// TIA Portal project "EXERCICE_IHM" (V16)

(* hardware
DEVICE "HMI_1"  KTP700 Basic PN
   slot 0: "HMI_1"  KTP700 Basic PN  6AV2 123-2GB03-0AX0  16.0.0.0
   slot 1: "HMI_RT_1"  KTP700 Basic PN  6AV2 123-2GB03-0AX0  16.0.0.0
   slot 5: "HMI_1.IE_CP_1"  PROFINET Interface  16.0.0.0
      slot 1: "Interface PROFINET_1"  PROFINET Interface
         slot 1: "Port_1"  Port
DEVICE "Station S7-1200_1"  S7-1200 Station
   slot 0: "Châssis_0"  S7-1200 Rack  Rack  V1.0
   slot 1: "PLC_1"  CPU 1214C AC/DC/Rly  6ES7 214-1BG40-0XB0  V4.4
*)

// ===== PLC "PLC_1"  CPU 1214C AC/DC/Rly =====

VAR_GLOBAL   // PLC tag table "Table de variables standard"
   "START" AT %I0.0 : Bool;
   "STOP" AT %I0.1 : Bool;
   "Moteur" AT %Q0.0 : Bool;
   "H1" AT %Q0.1 : Bool;
   "Clock_Byte" AT %MB0 : Byte;
   "Clock_10Hz" AT %M0.0 : Bool;
   "Clock_5Hz" AT %M0.1 : Bool;
   "Clock_2.5Hz" AT %M0.2 : Bool;
   "Clock_2Hz" AT %M0.3 : Bool;
   "Clock_1.25Hz" AT %M0.4 : Bool;
   "Clock_1Hz" AT %M0.5 : Bool;
   "Clock_0.625Hz" AT %M0.6 : Bool;
   "Clock_0.5Hz" AT %M0.7 : Bool;
   "HMI VENTILATEUR" AT %Q0.2 : Bool;
   "VENTILATEUR" AT %Q0.3 : Bool;
   "HMI MEMEUR" AT %Q0.4 : Bool;
END_VAR

ORGANIZATION_BLOCK "Main"   // OB1, LAD, ProgramCycle
TITLE = "Main Program Sweep (Cycle)"
{ S7_Optimized_Access := 'TRUE' }
VERSION : 0.1
   VAR_INPUT
      Initial_Call : Bool;   // Initial call of this OB
      Remanence : Bool;   // =True, if remanent data are available
   END_VAR
BEGIN

REGION Network 1
   // MOTEUR
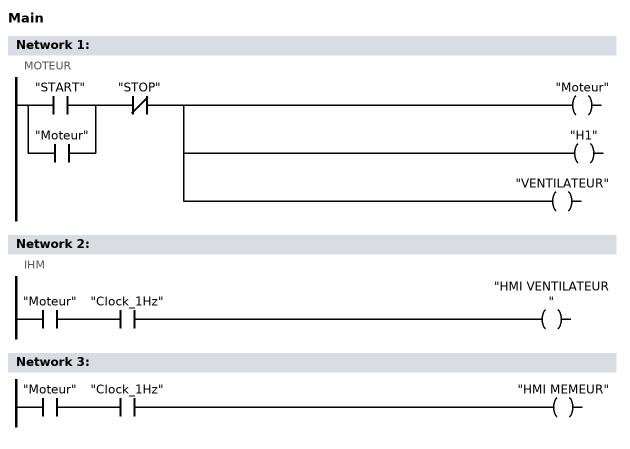
   RUNG wire#powerrail
      Contact( "START" )
      wire#w1
      I_Contact( "STOP" )
      wire#w2
      Coil( "Moteur" )
   END_RUNG
   RUNG wire#powerrail
      Contact( "Moteur" )
   END_RUNG wire#w1
   RUNG wire#w2
      Coil( "H1" )
   END_RUNG
   RUNG wire#w2
      Coil( "VENTILATEUR" )
   END_RUNG
   // the same network as SCL:
   "Moteur" := ("START" OR "Moteur") AND NOT "STOP";
   "H1" := "Moteur";
   "VENTILATEUR" := "Moteur";
END_REGION

REGION Network 2
   // IHM
   RUNG wire#powerrail
      Contact( "Moteur" )
      Contact( "Clock_1Hz" )
      Coil( "HMI VENTILATEUR" )
   END_RUNG
   // the same network as SCL:
   "HMI VENTILATEUR" := "Moteur" AND "Clock_1Hz";
END_REGION

REGION Network 3
   RUNG wire#powerrail
      Contact( "Moteur" )
      Contact( "Clock_1Hz" )
      Coil( "HMI MEMEUR" )
   END_RUNG
   // the same network as SCL:
   "HMI MEMEUR" := "Moteur" AND "Clock_1Hz";
END_REGION
END_ORGANIZATION_BLOCK

(* ===== HMI "HMI_RT_1" =====
system functions are stored by id; their names below are inferred from use
connection "HMI_Liaison_1": ETHERNET, SMART_S7_1200_OMS

HMI tags "Table de variables standard"
   "Numéro_vue_variable" : UInt, internal
   "START_IHM" : UInt, internal
   "START" : Bool = PLC START AT %I0.0, 100 ms
   "STOP" : Bool = PLC STOP AT %I0.1, 100 ms
   "HMI MEMEUR" : Bool = PLC "HMI MEMEUR" AT %Q0.4, 100 ms
   "H1" : Bool = PLC H1 AT %Q0.1, 100 ms
   "HMI VENTILATEUR" : Bool = PLC "HMI VENTILATEUR" AT %Q0.2, 100 ms

text list "Nom_vue_liste_textes": 1 'Vue racine'

Template "Modèle_1" 800x480
   Button "Quitter" at 714,429 size 71x50; TextOff 'Quitter'; PictureOff "ExitRuntime_KTP700_Basic_PN_TR"; PictureOn "ExitRuntime_KTP700_Basic_PN_TR"
      on Release: StopRuntime(0)
   Button "Template_Button" at 614,429 size 71x50; TextOff 'Text'
   Button "Template_Button_1" at 514,429 size 71x50; TextOff 'Text'
   Button "Template_Button_2" at 414,429 size 71x50; TextOff 'Text'
   Button "Template_Button_3" at 314,429 size 71x50; TextOff 'Text'
   Button "Template_Button_4" at 214,429 size 71x50; TextOff 'Text'
   Button "Template_Button_5" at 114,429 size 71x50; TextOff 'Text'
   Button "Vue initiale" at 14,429 size 71x50; TextOff 'Vue initiale'; PictureOff "NavigateHome_KTP700_Basic_PN_TR"; PictureOn "NavigateHome_KTP700_Basic_PN_TR"
      on Release: ActivateScreen("Vue racine", 0)
   SymbolicIOField "Vue_champ_ES_symbolique" at 93,9 size 600x33; TextOff '0'; TextOn '1'; TextList "Nom_vue_liste_textes"
      ProcessValue <- "Numéro_vue_variable"
      on Change: ActivateScreenByNumber("Numéro_vue_variable", 0)
   DateTimeField "HmiScreenItemData" at 695,25 size 105x25
   DateTimeField "HmiScreenItemData_1" at 695,0 size 105x25
   GraphicView "Logo" at 0,0 size 91x51; Picture "Logo de HMI_1"

screen "Vue racine" 800x480, template "Modèle_1"
   on GenerateScreen: SetTag("Numéro_vue_variable", 1)
   GraphicView "Vue de graphique_1" at 512,40 size 288x426; Picture "Graphique_1"
   GraphicView "Vue de graphique_7" at 573,155 size 178x178; Picture "Graphique_7"
      Visibility <- "HMI MEMEUR"
   TextField "HmiScreenItemData" at 0,0 size 800x45; Text 'MIXEUR HMI'
   Button "Bouton_1" at 41,116 size 96x32; TextOff 'START'
      on Press: SetBit("START")
   Button "Bouton_2" at 41,185 size 96x32; TextOff 'STOP'
      on Press: SetBit("STOP")
   GraphicView "Vue de graphique_2" at 369,284 size 134x134; Picture "Graphique_3"
      Visibility <- "HMI VENTILATEUR"
   GraphicView "Vue de graphique_3" at 360,32767 size 134x134; Picture "Graphique_3"
      Visibility <- "HMI VENTILATEUR"
   GraphicView "Vue de graphique_5" at 620,45 size 83x238; Picture "Graphique_5"
      Visibility <- "HMI MEMEUR"
   GraphicView "Vue de graphique_6" at 573,156 size 176x177; Picture "Graphique_6"
      Visibility <- "HMI MEMEUR"
   Circle "Cercle_1" at 442,104 size 38x38
      Appearance <- "H1"
   GraphicView "Vue de graphique_4" at 621,46 size 83x238; Picture "Graphique_4"
      Visibility <- "HMI MEMEUR"
*)